(* Logix 5000 project; controller TFF vendor 1 type 14 code 107 rev 34.11; software revision 34.03; part 23 of 36 *)
(* tags used below, declared in another part *)
   Address : DINT;   // Temp Address
   Address2 : DINT;   // Temp Address
   FeedPump_PID_Settings : INT;   // Index
   Index : DINT;   // Index
   ONS_PID02 : BOOL;
   SCL : SCALE;   // Scale Instruction
   AnalogOutput : AnalogOutput[25];   // Analog Output Array
   AnalogPoint : AnalogInput[50];   // Analog Input Array
   ControlLoop : ControlLoop[20];   // Control Loop Array
   ControlLoop_FeedPump : ALIAS FOR ControlLoop[1];   // Feed Pump Control Loop
   ControlLoop_PCV001 : ALIAS FOR ControlLoop[3];   // PCV001 Control Loop
   ControlLoop_PCV001_5ms : ALIAS FOR ControlLoop[4];   // PCV001 Control Loop
   ControlLoop_PCV001_RAMP_OUT : REAL;   // Ramp Output
   ControlLoop_PCV101 : ALIAS FOR ControlLoop[5];   // PCV101 Control Loop
   Mixer : Mixer;   // Mixer config. structure
   PCV001 : ALIAS FOR AnalogPoint[3];   // Retentate Pressure Control Valve Position
   PCV001_Control : PCV_Control;   // PCV001 Control UDT
   PumpRunStatus : DINT;   // Pumps Run Status (1 = At least one pump running , 0 = no pump running)
   SIC003 : ALIAS FOR Drive[3];   // Mixer
   SIC003_AO : ALIAS FOR AnalogOutput[4];   // Mixer Speed Setpoint
   SysControl : SysControl;   // General system status and command
   WI001 : ALIAS FOR AnalogPoint[15];   // Feed Bag Weight
(* Process, continued *)

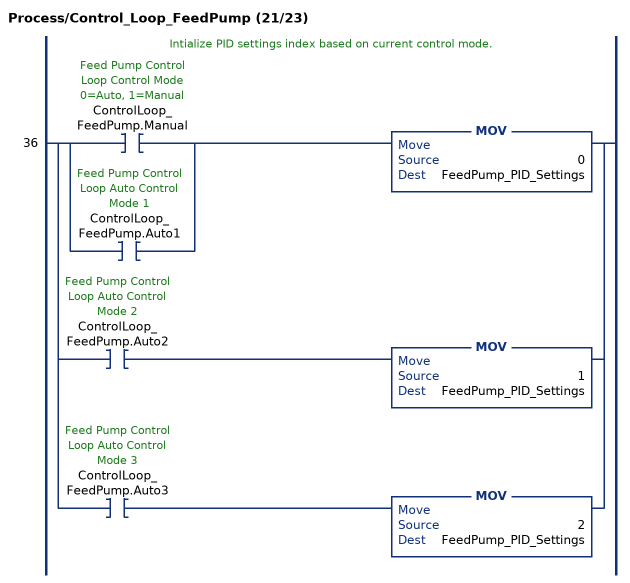
   [picture p189: Process/Control_Loop_FeedPump rungs 36-36]
   // Intialize PID settings index based on current control mode.
   36: [[XIC(ControlLoop_FeedPump.Manual) ,XIC(ControlLoop_FeedPump.Auto1) ] MOV(0,FeedPump_PID_Settings) ,XIC(ControlLoop_FeedPump.Auto2) MOV(1,FeedPump_PID_Settings) ,XIC(ControlLoop_FeedPump.Auto3) MOV(2,FeedPump_PID_Settings) ];
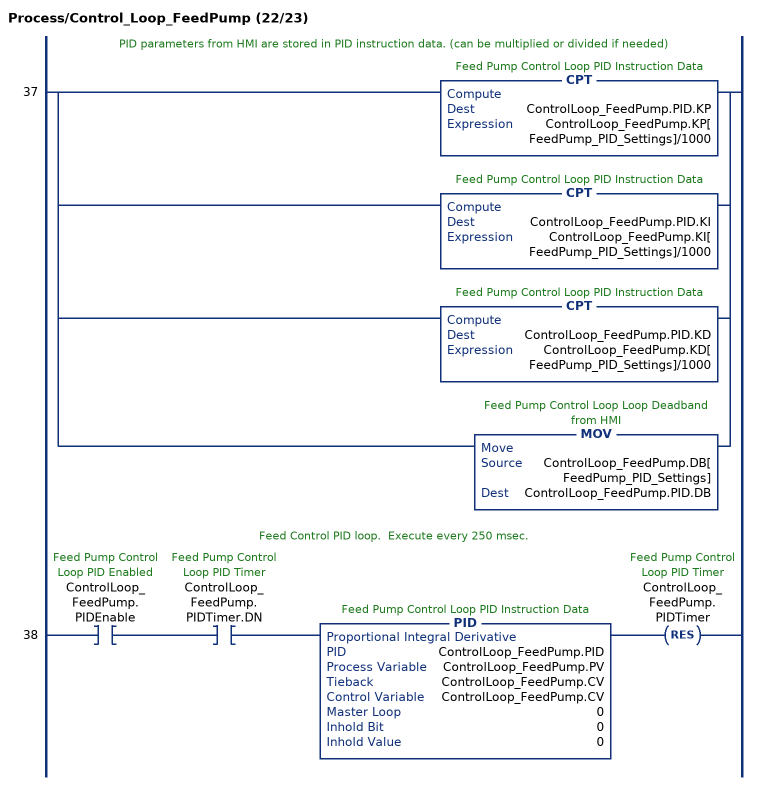
   // PID parameters from HMI are stored in PID instruction data. (can be multiplied or divided if needed)
   37: [CPT(ControlLoop_FeedPump.PID.KP,ControlLoop_FeedPump.KP[FeedPump_PID_Settings]/1000) ,CPT(ControlLoop_FeedPump.PID.KI,ControlLoop_FeedPump.KI[FeedPump_PID_Settings]/1000) ,CPT(ControlLoop_FeedPump.PID.KD,ControlLoop_FeedPump.KD[FeedPump_PID_Settings]/1000) ,MOV(ControlLoop_FeedPump.DB[FeedPump_PID_Settings],ControlLoop_FeedPump.PID.DB) ];
   // Feed Control PID loop.  Execute every 250 msec.
   38: XIC(ControlLoop_FeedPump.PIDEnable)XIC(ControlLoop_FeedPump.PIDTimer.DN)PID(ControlLoop_FeedPump.PID,ControlLoop_FeedPump.PV,ControlLoop_FeedPump.CV,ControlLoop_FeedPump.CV,0,0,0)RES(ControlLoop_FeedPump.PIDTimer);
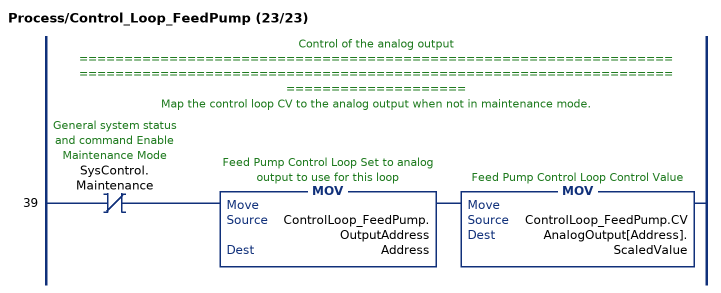
   // Control of the analog output
   // ========================================================================================================================================================
   // Map the control loop CV to the analog output when not in maintenance mode.
   39: XIO(SysControl.Maintenance)MOV(ControlLoop_FeedPump.OutputAddress,Address)MOV(ControlLoop_FeedPump.CV,AnalogOutput[Address].ScaledValue);
END_ROUTINE

ROUTINE Control_Loop_Mixer   (* ladder *)
// Agitator Control Routine
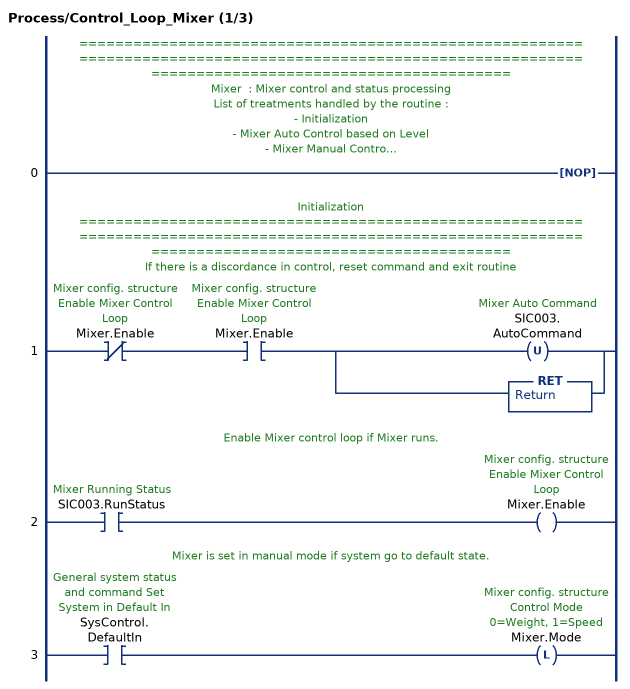
   // ========================================================================================================================================================
   //                                                                                                    Mixer  : Mixer control and status processing
   //                                                     List of treatments handled by the routine :
   //                                                          - Initialization
   //                                                          - Mixer Auto Control based on Level
   //                                                          - Mixer Manual Control
   //                                                     -----------------------------------------------------------------------------------------------------------------------------------------------------
   //                                                     History
   //                                                          2019-AUG-13 - Actemium - B. Roch - Initial version for Candidate Release 3.00.00.00.a
   // ========================================================================================================================================================
   0: NOP();
   // Initialization
   // ========================================================================================================================================================
   // If there is a discordance in control, reset command and exit routine
   1: XIO(Mixer.Enable)XIC(Mixer.Enable)[OTU(SIC003.AutoCommand) ,RET() ];
   // Enable Mixer control loop if Mixer runs.
   2: XIC(SIC003.RunStatus)OTE(Mixer.Enable);
   // Mixer is set in manual mode if system go to default state.
   3: XIC(SysControl.DefaultIn)OTL(Mixer.Mode);
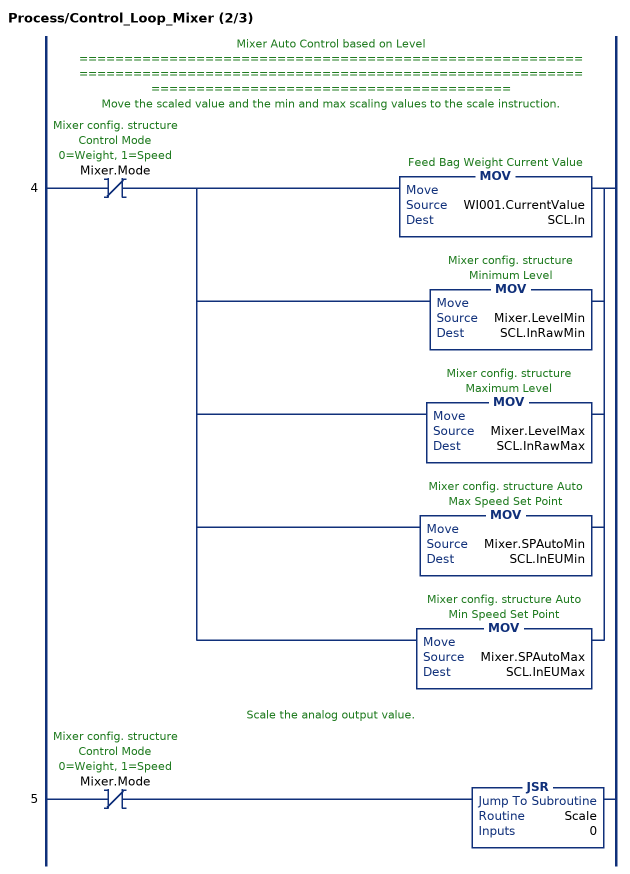
   // Mixer Auto Control based on Level
   // ========================================================================================================================================================
   // Move the scaled value and the min and max scaling values to the scale instruction.
   4: XIO(Mixer.Mode)[MOV(WI001.CurrentValue,SCL.In) ,MOV(Mixer.LevelMin,SCL.InRawMin) ,MOV(Mixer.LevelMax,SCL.InRawMax) ,MOV(Mixer.SPAutoMin,SCL.InEUMin) ,MOV(Mixer.SPAutoMax,SCL.InEUMax) ];
   // Scale the analog output value.
   5: XIO(Mixer.Mode)JSR(Scale,0);
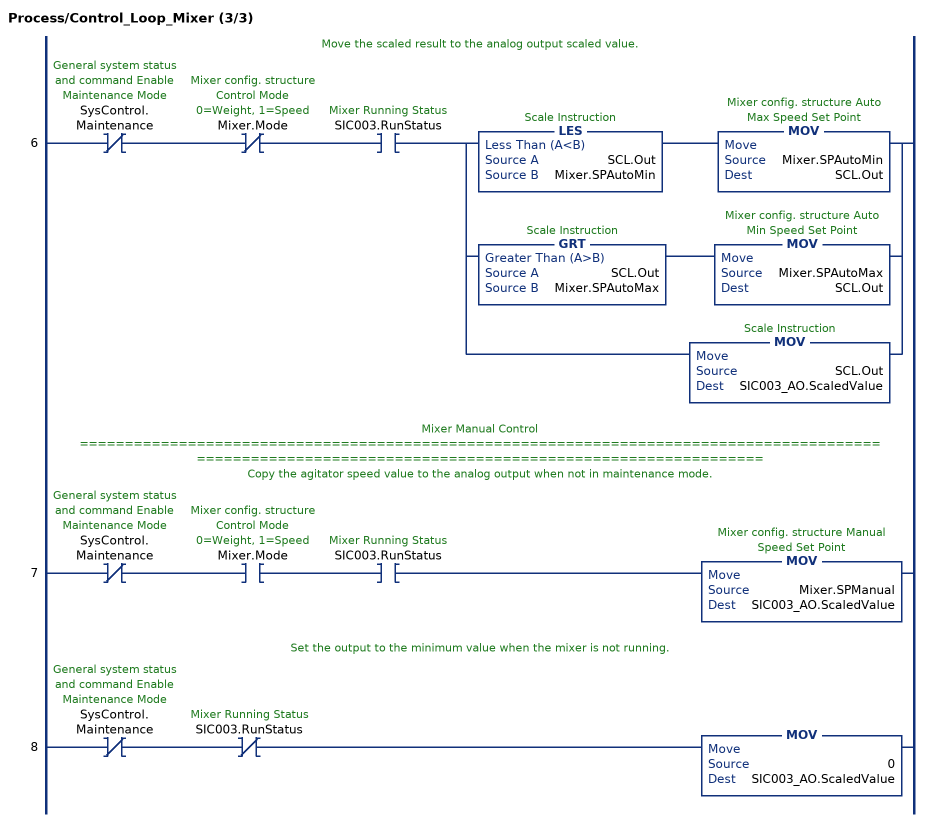
   // Move the scaled result to the analog output scaled value.
   6: XIO(SysControl.Maintenance)XIO(Mixer.Mode)XIC(SIC003.RunStatus)[LES(SCL.Out,Mixer.SPAutoMin) MOV(Mixer.SPAutoMin,SCL.Out) ,GRT(SCL.Out,Mixer.SPAutoMax) MOV(Mixer.SPAutoMax,SCL.Out) ,MOV(SCL.Out,SIC003_AO.ScaledValue) ];
   // Mixer Manual Control
   // ========================================================================================================================================================
   // Copy the agitator speed value to the analog output when not in maintenance mode.
   7: XIO(SysControl.Maintenance)XIC(Mixer.Mode)XIC(SIC003.RunStatus)MOV(Mixer.SPManual,SIC003_AO.ScaledValue);
   // Set the output to the minimum value when the mixer is not running.
   8: XIO(SysControl.Maintenance)XIO(SIC003.RunStatus)MOV(0,SIC003_AO.ScaledValue);
END_ROUTINE

ROUTINE Control_Loop_PCV001   (* ladder *)
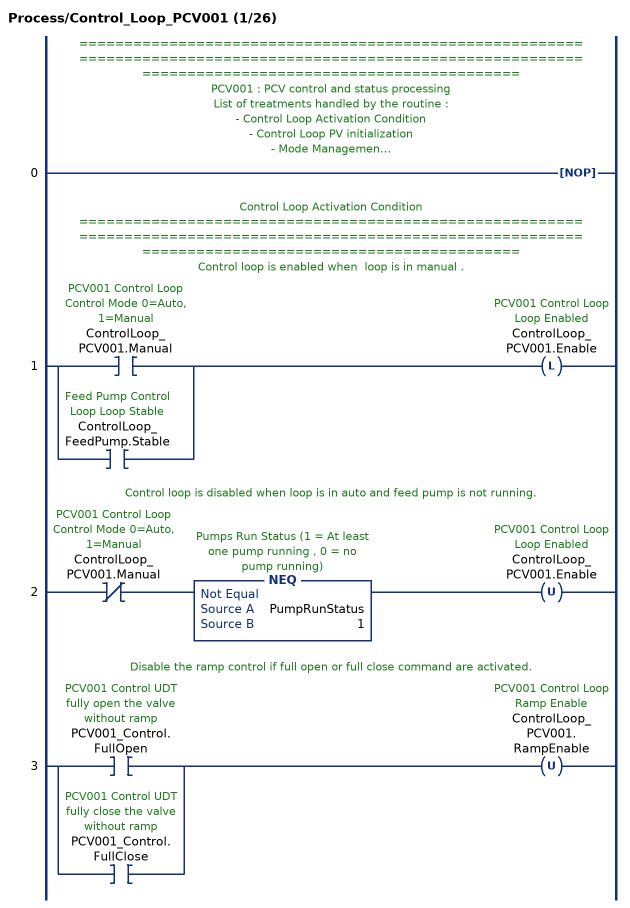
   // ==========================================================================================================================================================
   //                                                  PCV001 : PCV control and status processing
   //                                                     List of treatments handled by the routine :
   //                                                          - Control Loop Activation Condition
   //                                                  - Control Loop PV initialization
   //                                                - Mode Management
   //                                                        - Control Loop Setpoint management
   //                                                        - Control Loop deadband calculation
   //                                                          - Management of ramping control
   //                                                          - Control Loop Stability control
   //                                                          - Full Open - Full Close processing
   //                                                          - Management of PID instruction
   //                                                          - Control of the analog output
   //                                                     -----------------------------------------------------------------------------------------------------------------------------------------------------
   //                                                     History
   //                                2019-SEP-26 - Actemium - B. Roch - Initial version for Candidate Release 3.00.00.00.c                               2020-SEP-14 - Merck - Q. Spindler - Modifications for Candidate Release 3.00.00.01.a
   //                                                        - on rung 17, disable DBOK if control loop is not enabled or in manual
   // 	2021-APR-19 - DAVIDSON- Ch. ARBOGAST - Modifications for Candidate Release 3.01.00.00.a
   // 	- on rung 4, line 1, replace "ControlLoop[3].Manual OR ControlLoop[3].Auto1" by
   // 			 "NOT ControlLoop[3].Auto2 AND NOT ControlLoop[3].Auto3"
   // ==========================================================================================================================================================
   0: NOP();
   // Control Loop Activation Condition
   // ==========================================================================================================================================================
   // Control loop is enabled when  loop is in manual .
   1: [XIC(ControlLoop_PCV001.Manual) ,XIC(ControlLoop_FeedPump.Stable) ]OTL(ControlLoop_PCV001.Enable);
   // Control loop is disabled when loop is in auto and feed pump is not running.
   2: XIO(ControlLoop_PCV001.Manual)NEQ(PumpRunStatus,1)OTU(ControlLoop_PCV001.Enable);
   // Disable the ramp control if full open or full close command are activated.
   3: [XIC(PCV001_Control.FullOpen) ,XIC(PCV001_Control.FullClose) ]OTU(ControlLoop_PCV001.RampEnable);
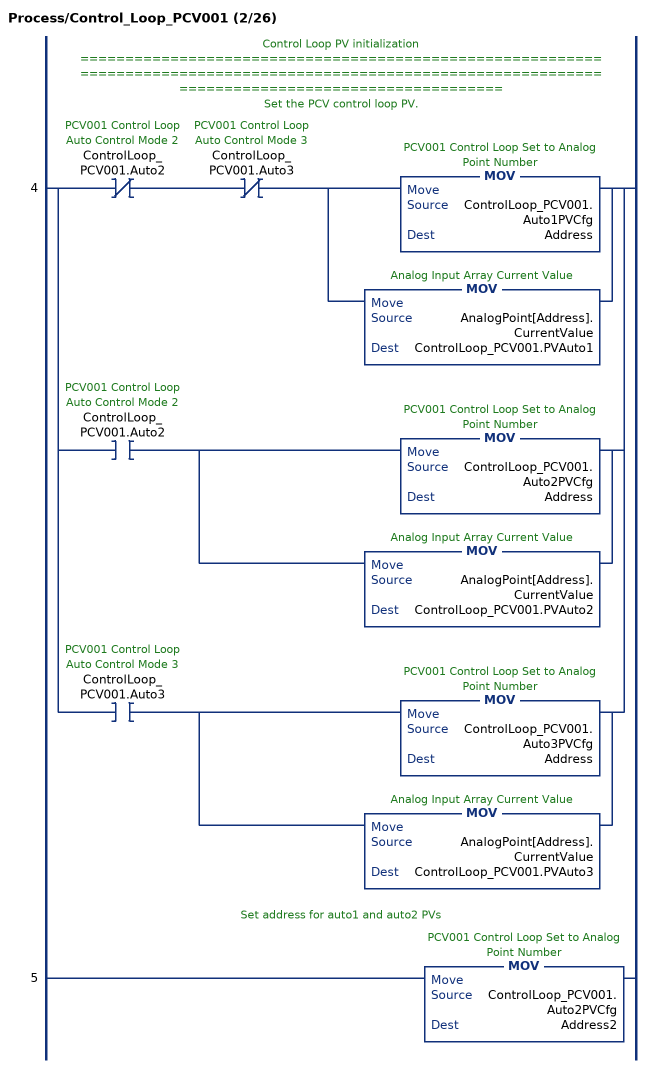
   // Control Loop PV initialization
   // ========================================================================================================================================================
   // Set the PCV control loop PV.
   4: [[XIO(ControlLoop_PCV001.Auto2) XIO(ControlLoop_PCV001.Auto3) [MOV(ControlLoop_PCV001.Auto1PVCfg,Address) ,MOV(AnalogPoint[Address].CurrentValue,ControlLoop_PCV001.PVAuto1) ] ,XIC(ControlLoop_PCV001.Auto2) [MOV(ControlLoop_PCV001.Auto2PVCfg,Address) ,MOV(AnalogPoint[Address].CurrentValue,ControlLoop_PCV001.PVAuto2) ] ] ,XIC(ControlLoop_PCV001.Auto3) [MOV(ControlLoop_PCV001.Auto3PVCfg,Address) ,MOV(AnalogPoint[Address].CurrentValue,ControlLoop_PCV001.PVAuto3) ] ];
   // Set address for auto1 and auto2 PVs
   5: MOV(ControlLoop_PCV001.Auto2PVCfg,Address2);
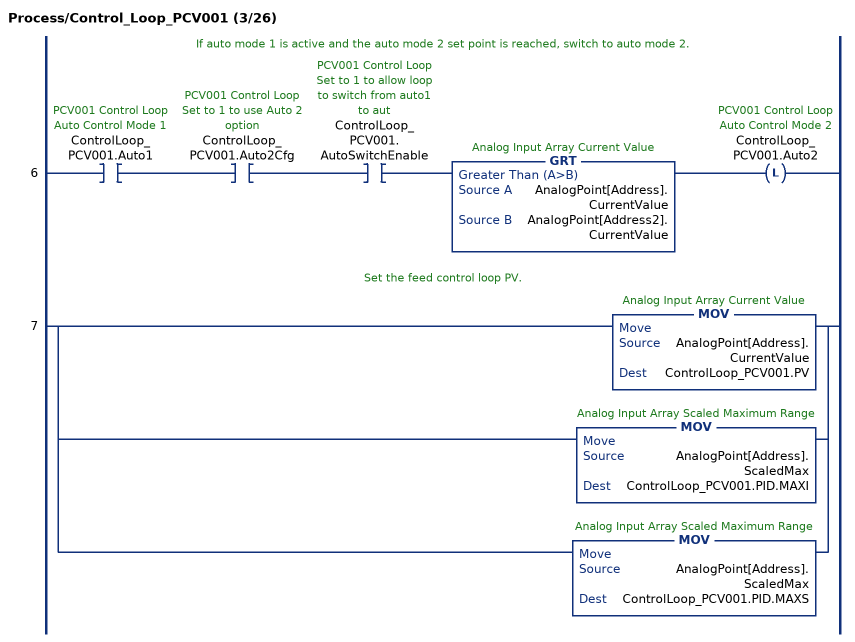
   // If auto mode 1 is active and the auto mode 2 set point is reached, switch to auto mode 2.
   6: XIC(ControlLoop_PCV001.Auto1)XIC(ControlLoop_PCV001.Auto2Cfg)XIC(ControlLoop_PCV001.AutoSwitchEnable)GRT(AnalogPoint[Address].CurrentValue,AnalogPoint[Address2].CurrentValue)OTL(ControlLoop_PCV001.Auto2);
   // Set the feed control loop PV.
   7: [MOV(AnalogPoint[Address].CurrentValue,ControlLoop_PCV001.PV) ,MOV(AnalogPoint[Address].ScaledMax,ControlLoop_PCV001.PID.MAXI) ,MOV(AnalogPoint[Address].ScaledMax,ControlLoop_PCV001.PID.MAXS) ];
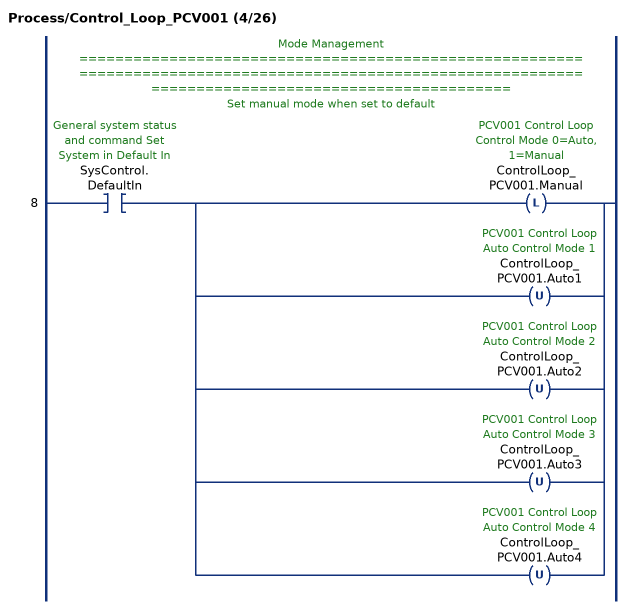
   // Mode Management
   // ========================================================================================================================================================
   // Set manual mode when set to default
   8: XIC(SysControl.DefaultIn)[OTL(ControlLoop_PCV001.Manual) ,OTU(ControlLoop_PCV001.Auto1) ,OTU(ControlLoop_PCV001.Auto2) ,OTU(ControlLoop_PCV001.Auto3) ,OTU(ControlLoop_PCV001.Auto4) ];
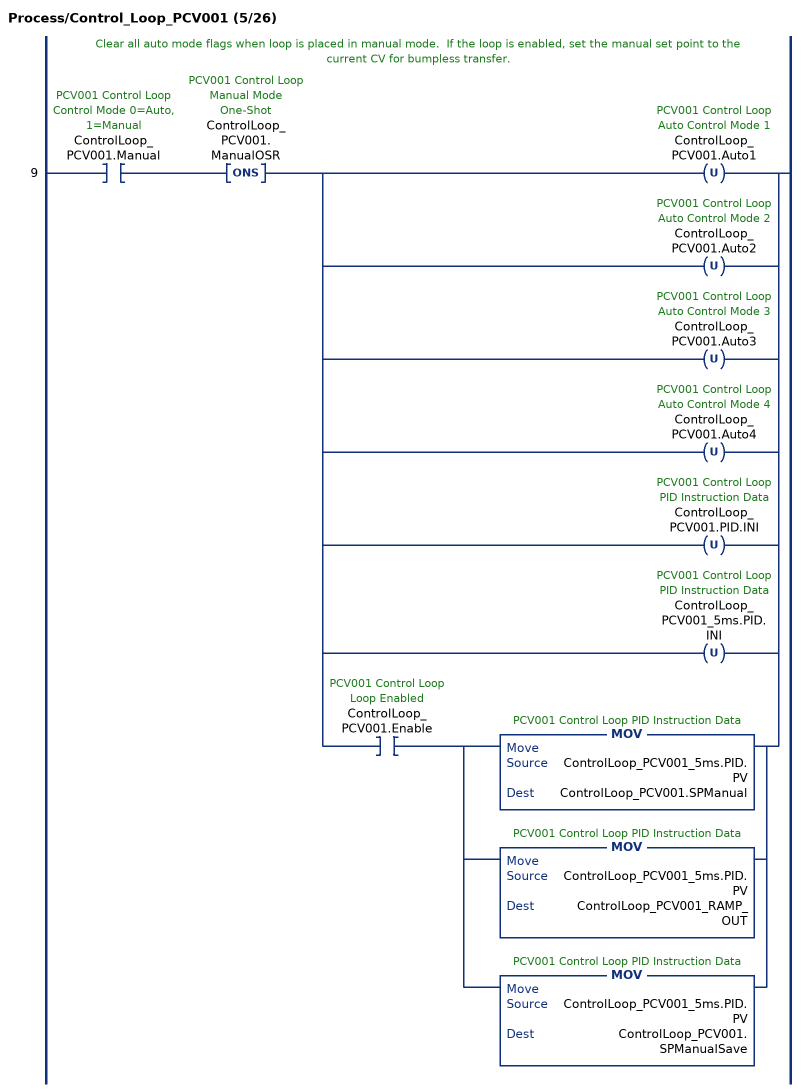
   // Clear all auto mode flags when loop is placed in manual mode.  If the loop is enabled, set the manual set point to the current CV for bumpless transfer.
   9: XIC(ControlLoop_PCV001.Manual)ONS(ControlLoop_PCV001.ManualOSR)[OTU(ControlLoop_PCV001.Auto1) ,OTU(ControlLoop_PCV001.Auto2) ,OTU(ControlLoop_PCV001.Auto3) ,OTU(ControlLoop_PCV001.Auto4) ,OTU(ControlLoop_PCV001.PID.INI) ,OTU(ControlLoop_PCV001_5ms.PID.INI) ,XIC(ControlLoop_PCV001.Enable) [MOV(ControlLoop_PCV001_5ms.PID.PV,ControlLoop_PCV001.SPManual) ,MOV(ControlLoop_PCV001_5ms.PID.PV,ControlLoop_PCV001_RAMP_OUT) ,MOV(ControlLoop_PCV001_5ms.PID.PV,ControlLoop_PCV001.SPManualSave) ] ];
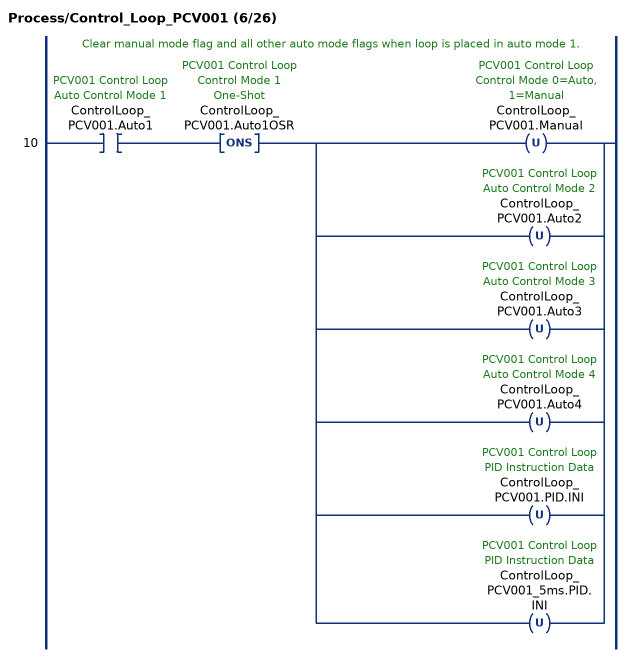
   // Clear manual mode flag and all other auto mode flags when loop is placed in auto mode 1.
   10: XIC(ControlLoop_PCV001.Auto1)ONS(ControlLoop_PCV001.Auto1OSR)[OTU(ControlLoop_PCV001.Manual) ,OTU(ControlLoop_PCV001.Auto2) ,OTU(ControlLoop_PCV001.Auto3) ,OTU(ControlLoop_PCV001.Auto4) ,OTU(ControlLoop_PCV001.PID.INI) ,OTU(ControlLoop_PCV001_5ms.PID.INI) ];
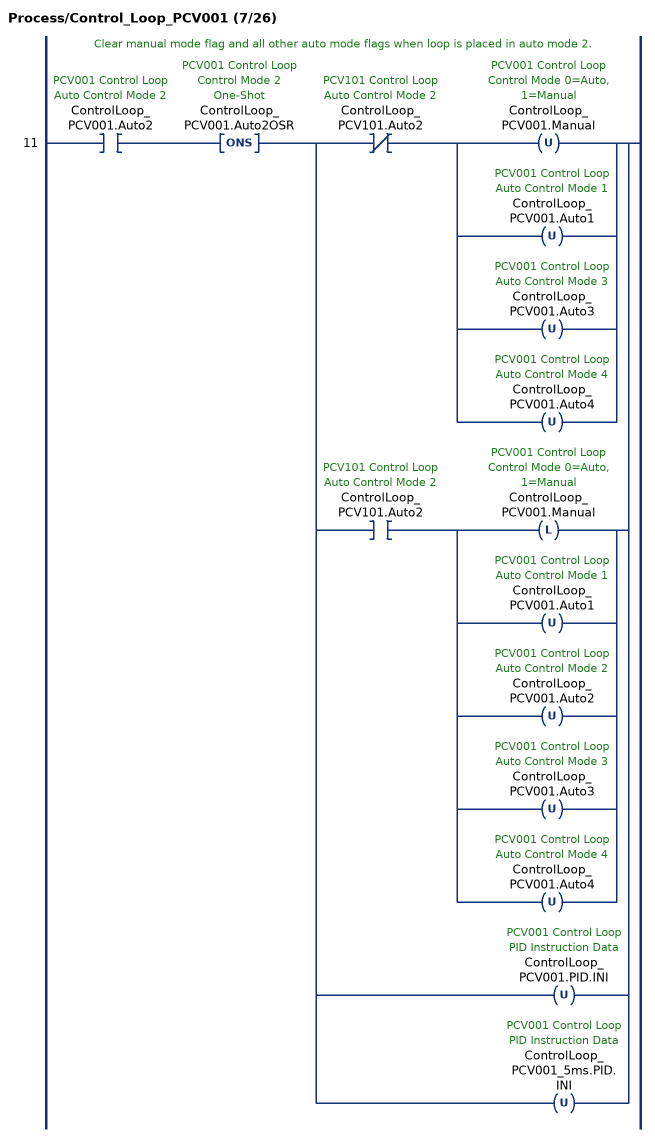
   // Clear manual mode flag and all other auto mode flags when loop is placed in auto mode 2.
   11: XIC(ControlLoop_PCV001.Auto2)ONS(ControlLoop_PCV001.Auto2OSR)[XIO(ControlLoop_PCV101.Auto2) [OTU(ControlLoop_PCV001.Manual) ,OTU(ControlLoop_PCV001.Auto1) ,OTU(ControlLoop_PCV001.Auto3) ,OTU(ControlLoop_PCV001.Auto4) ] ,XIC(ControlLoop_PCV101.Auto2) [OTL(ControlLoop_PCV001.Manual) ,OTU(ControlLoop_PCV001.Auto1) ,OTU(ControlLoop_PCV001.Auto2) ,OTU(ControlLoop_PCV001.Auto3) ,OTU(ControlLoop_PCV001.Auto4) ] ,OTU(ControlLoop_PCV001.PID.INI) ,OTU(ControlLoop_PCV001_5ms.PID.INI) ];
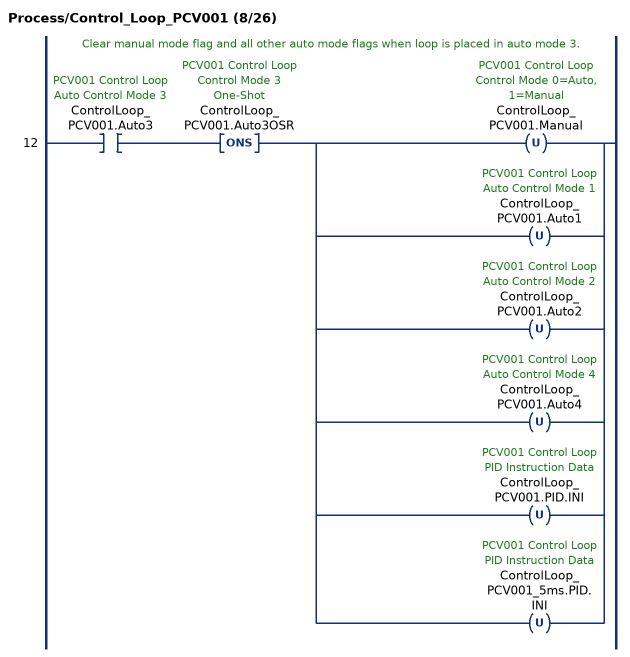
   // Clear manual mode flag and all other auto mode flags when loop is placed in auto mode 3.
   12: XIC(ControlLoop_PCV001.Auto3)ONS(ControlLoop_PCV001.Auto3OSR)[OTU(ControlLoop_PCV001.Manual) ,OTU(ControlLoop_PCV001.Auto1) ,OTU(ControlLoop_PCV001.Auto2) ,OTU(ControlLoop_PCV001.Auto4) ,OTU(ControlLoop_PCV001.PID.INI) ,OTU(ControlLoop_PCV001_5ms.PID.INI) ];
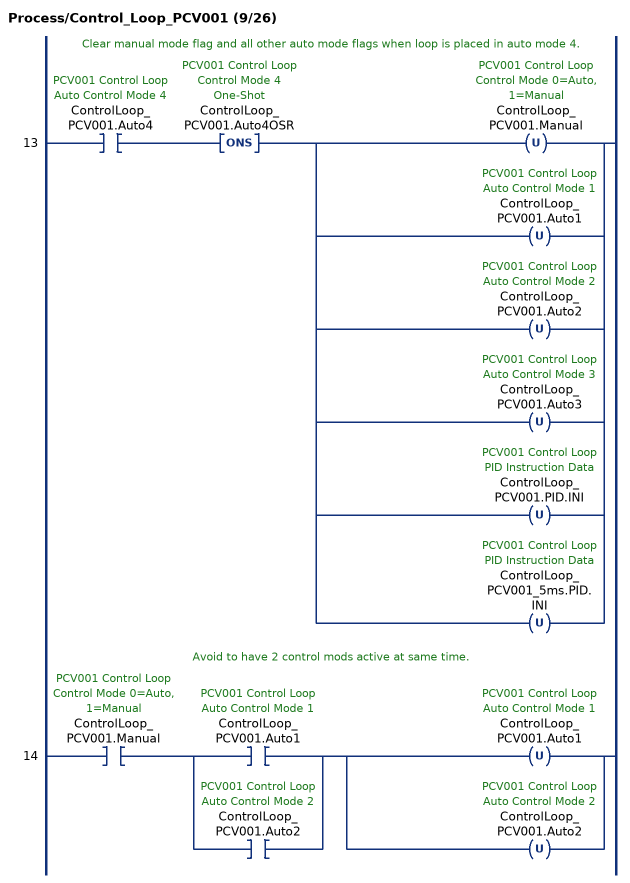
   // Clear manual mode flag and all other auto mode flags when loop is placed in auto mode 4.
   13: XIC(ControlLoop_PCV001.Auto4)ONS(ControlLoop_PCV001.Auto4OSR)[OTU(ControlLoop_PCV001.Manual) ,OTU(ControlLoop_PCV001.Auto1) ,OTU(ControlLoop_PCV001.Auto2) ,OTU(ControlLoop_PCV001.Auto3) ,OTU(ControlLoop_PCV001.PID.INI) ,OTU(ControlLoop_PCV001_5ms.PID.INI) ];
   // Avoid to have 2 control mods active at same time.
   14: XIC(ControlLoop_PCV001.Manual)[XIC(ControlLoop_PCV001.Auto1) ,XIC(ControlLoop_PCV001.Auto2) ][OTU(ControlLoop_PCV001.Auto1) ,OTU(ControlLoop_PCV001.Auto2) ];
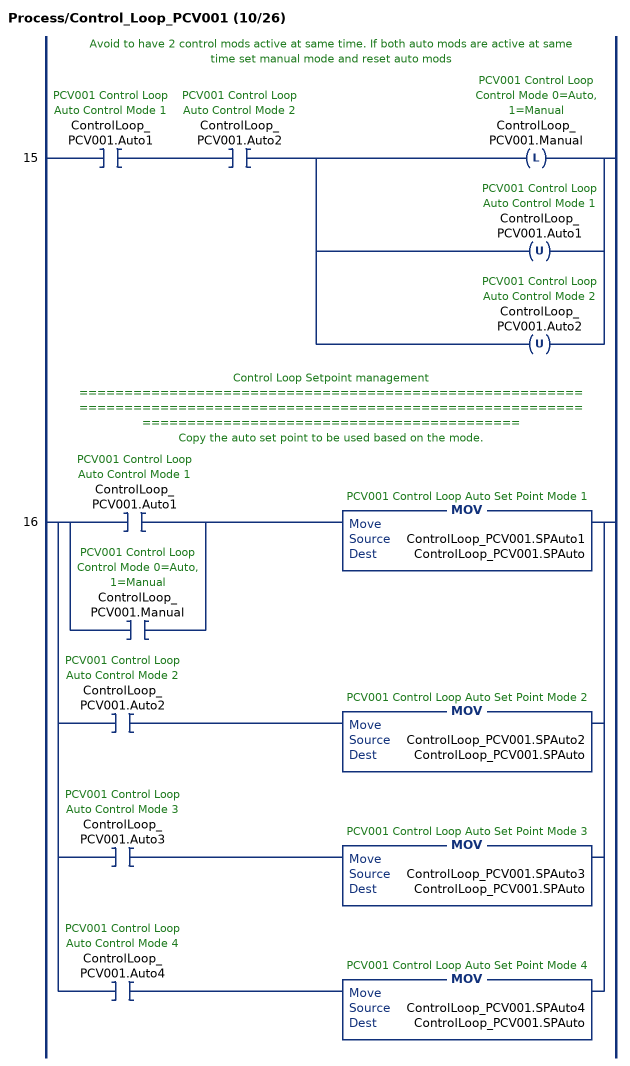
   // Avoid to have 2 control mods active at same time. If both auto mods are active at same time set manual mode and reset auto mods
   15: XIC(ControlLoop_PCV001.Auto1)XIC(ControlLoop_PCV001.Auto2)[OTL(ControlLoop_PCV001.Manual) ,OTU(ControlLoop_PCV001.Auto1) ,OTU(ControlLoop_PCV001.Auto2) ];
   // Control Loop Setpoint management
   // ==========================================================================================================================================================
   // Copy the auto set point to be used based on the mode.
   16: [[XIC(ControlLoop_PCV001.Auto1) ,XIC(ControlLoop_PCV001.Manual) ] MOV(ControlLoop_PCV001.SPAuto1,ControlLoop_PCV001.SPAuto) ,XIC(ControlLoop_PCV001.Auto2) MOV(ControlLoop_PCV001.SPAuto2,ControlLoop_PCV001.SPAuto) ,XIC(ControlLoop_PCV001.Auto3) MOV(ControlLoop_PCV001.SPAuto3,ControlLoop_PCV001.SPAuto) ,XIC(ControlLoop_PCV001.Auto4) MOV(ControlLoop_PCV001.SPAuto4,ControlLoop_PCV001.SPAuto) ];
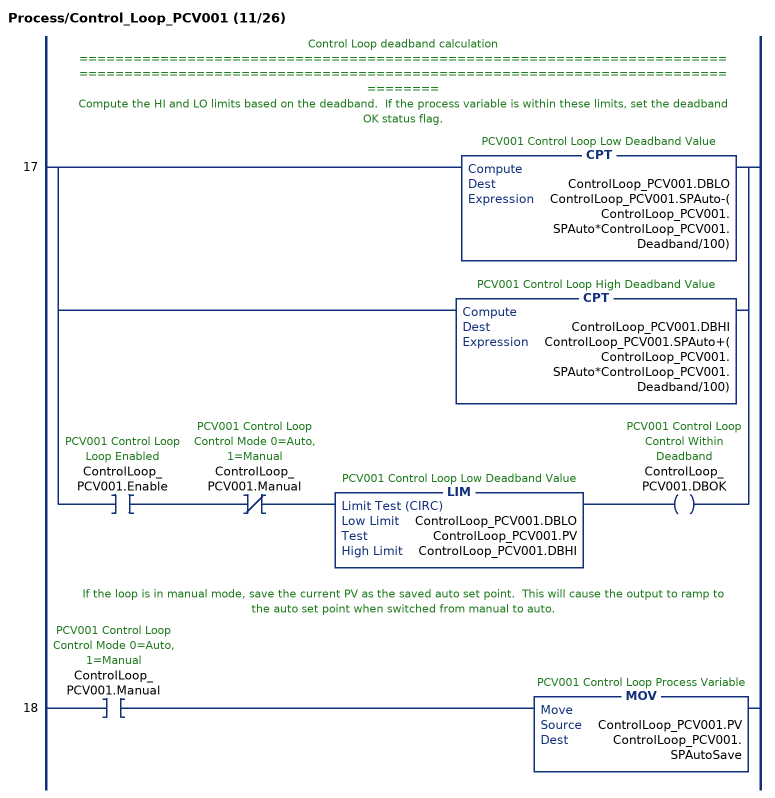
   // Control Loop deadband calculation
   // ========================================================================================================================================================
   // Compute the HI and LO limits based on the deadband.  If the process variable is within these limits, set the deadband OK status flag.
   17: [CPT(ControlLoop_PCV001.DBLO,ControlLoop_PCV001.SPAuto-(ControlLoop_PCV001.SPAuto*ControlLoop_PCV001.Deadband/100)) ,CPT(ControlLoop_PCV001.DBHI,ControlLoop_PCV001.SPAuto+(ControlLoop_PCV001.SPAuto*ControlLoop_PCV001.Deadband/100)) ,XIC(ControlLoop_PCV001.Enable) XIO(ControlLoop_PCV001.Manual) LIM(ControlLoop_PCV001.DBLO,ControlLoop_PCV001.PV,ControlLoop_PCV001.DBHI) OTE(ControlLoop_PCV001.DBOK) ];
   // If the loop is in manual mode, save the current PV as the saved auto set point.  This will cause the output to ramp to the auto set point when switched from manual to auto.
   18: XIC(ControlLoop_PCV001.Manual)MOV(ControlLoop_PCV001.PV,ControlLoop_PCV001.SPAutoSave);
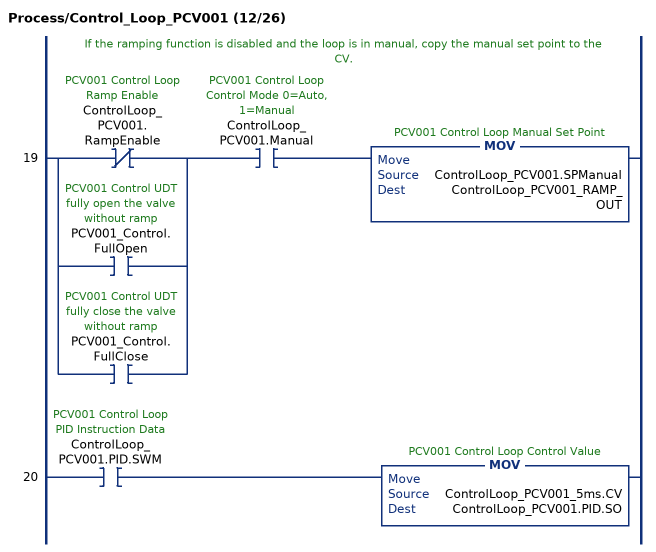
   // If the ramping function is disabled and the loop is in manual, copy the manual set point to the CV.
   19: [XIO(ControlLoop_PCV001.RampEnable) ,XIC(PCV001_Control.FullOpen) ,XIC(PCV001_Control.FullClose) ]XIC(ControlLoop_PCV001.Manual)MOV(ControlLoop_PCV001.SPManual,ControlLoop_PCV001_RAMP_OUT);
   20: XIC(ControlLoop_PCV001.PID.SWM)MOV(ControlLoop_PCV001_5ms.CV,ControlLoop_PCV001.PID.SO);
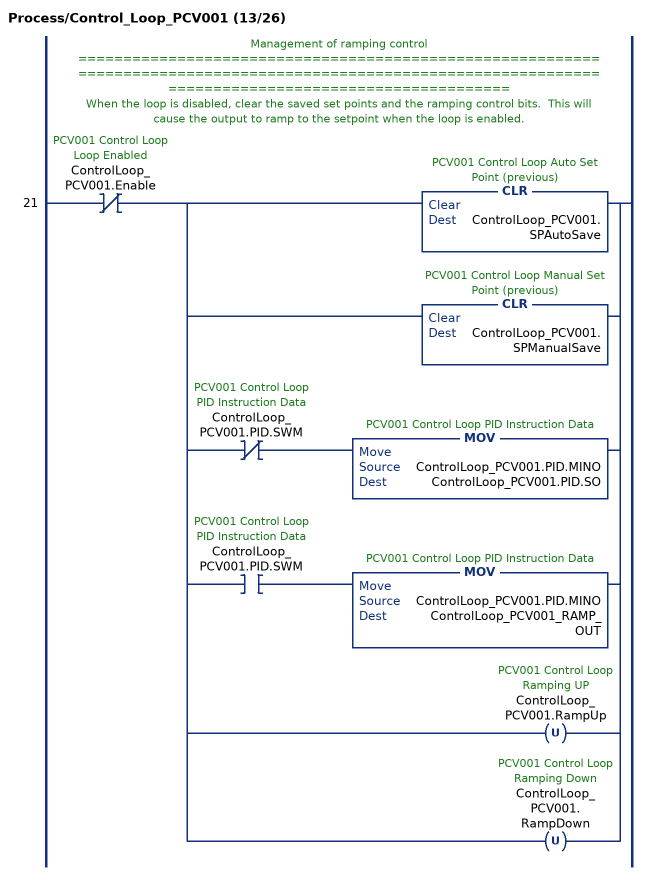
   // Management of ramping control
   // ==========================================================================================================================================================
   // When the loop is disabled, clear the saved set points and the ramping control bits.  This will cause the output to ramp to the setpoint when the loop is enabled.
   21: XIO(ControlLoop_PCV001.Enable)[CLR(ControlLoop_PCV001.SPAutoSave) ,CLR(ControlLoop_PCV001.SPManualSave) ,XIO(ControlLoop_PCV001.PID.SWM) MOV(ControlLoop_PCV001.PID.MINO,ControlLoop_PCV001.PID.SO) ,XIC(ControlLoop_PCV001.PID.SWM) MOV(ControlLoop_PCV001.PID.MINO,ControlLoop_PCV001_RAMP_OUT) ,OTU(ControlLoop_PCV001.RampUp) ,OTU(ControlLoop_PCV001.RampDown) ];
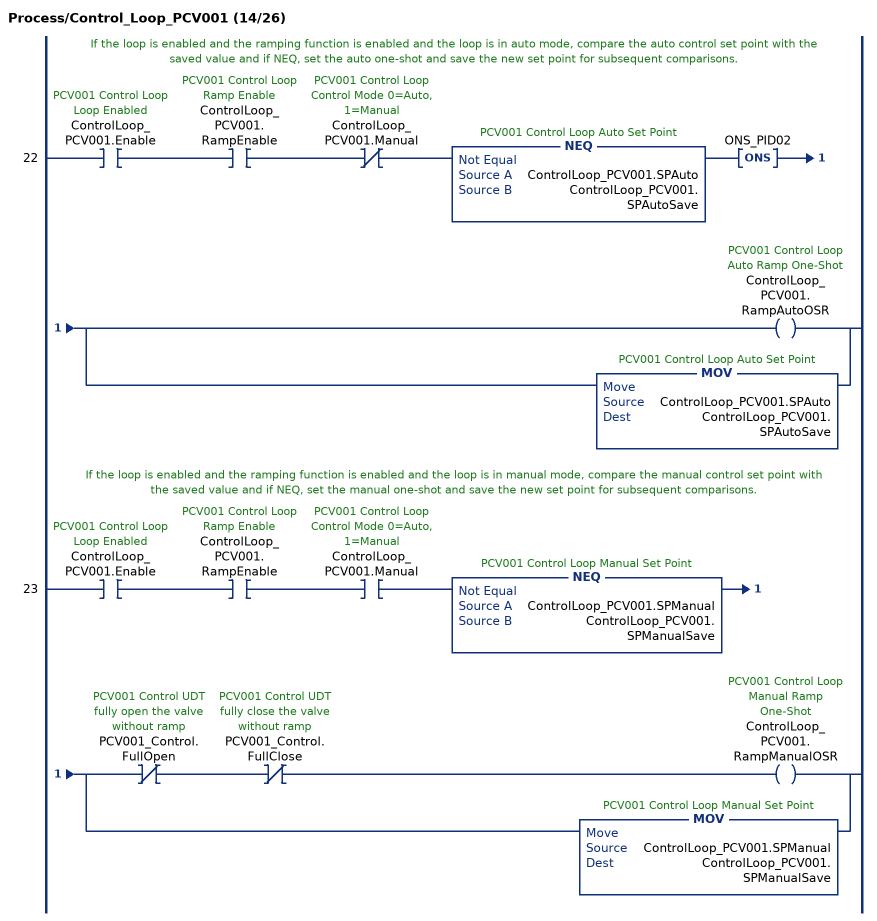
   // If the loop is enabled and the ramping function is enabled and the loop is in auto mode, compare the auto control set point with the saved value and if NEQ, set the auto one-shot and save the new set point for subsequent comparisons.
   22: XIC(ControlLoop_PCV001.Enable)XIC(ControlLoop_PCV001.RampEnable)XIO(ControlLoop_PCV001.Manual)NEQ(ControlLoop_PCV001.SPAuto,ControlLoop_PCV001.SPAutoSave)ONS(ONS_PID02)[OTE(ControlLoop_PCV001.RampAutoOSR) ,MOV(ControlLoop_PCV001.SPAuto,ControlLoop_PCV001.SPAutoSave) ];
   // If the loop is enabled and the ramping function is enabled and the loop is in manual mode, compare the manual control set point with the saved value and if NEQ, set the manual one-shot and save the new set point for subsequent comparisons.
   23: XIC(ControlLoop_PCV001.Enable)XIC(ControlLoop_PCV001.RampEnable)XIC(ControlLoop_PCV001.Manual)NEQ(ControlLoop_PCV001.SPManual,ControlLoop_PCV001.SPManualSave)[XIO(PCV001_Control.FullOpen) XIO(PCV001_Control.FullClose) OTE(ControlLoop_PCV001.RampManualOSR) ,MOV(ControlLoop_PCV001.SPManual,ControlLoop_PCV001.SPManualSave) ];
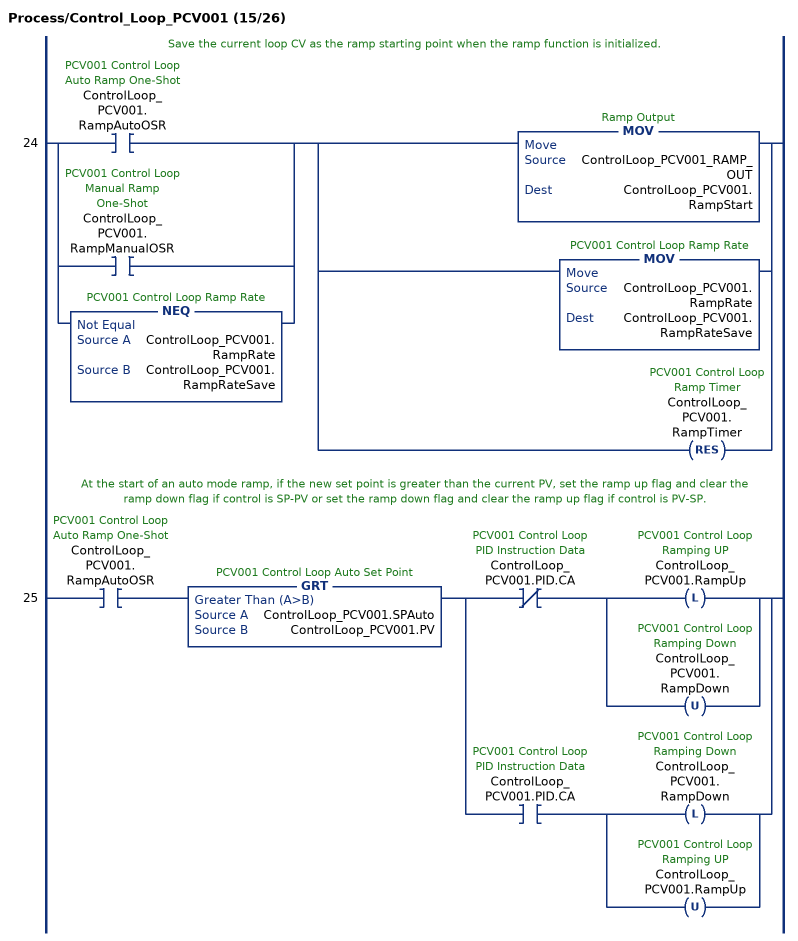
   // Save the current loop CV as the ramp starting point when the ramp function is initialized.
   24: [XIC(ControlLoop_PCV001.RampAutoOSR) ,XIC(ControlLoop_PCV001.RampManualOSR) ,NEQ(ControlLoop_PCV001.RampRate,ControlLoop_PCV001.RampRateSave) ][MOV(ControlLoop_PCV001_RAMP_OUT,ControlLoop_PCV001.RampStart) ,MOV(ControlLoop_PCV001.RampRate,ControlLoop_PCV001.RampRateSave) ,RES(ControlLoop_PCV001.RampTimer) ];
   // At the start of an auto mode ramp, if the new set point is greater than the current PV, set the ramp up flag and clear the ramp down flag if control is SP-PV or set the ramp down flag and clear the ramp up flag if control is PV-SP.
   25: XIC(ControlLoop_PCV001.RampAutoOSR)GRT(ControlLoop_PCV001.SPAuto,ControlLoop_PCV001.PV)[XIO(ControlLoop_PCV001.PID.CA) [OTL(ControlLoop_PCV001.RampUp) ,OTU(ControlLoop_PCV001.RampDown) ] ,XIC(ControlLoop_PCV001.PID.CA) [OTL(ControlLoop_PCV001.RampDown) ,OTU(ControlLoop_PCV001.RampUp) ] ];
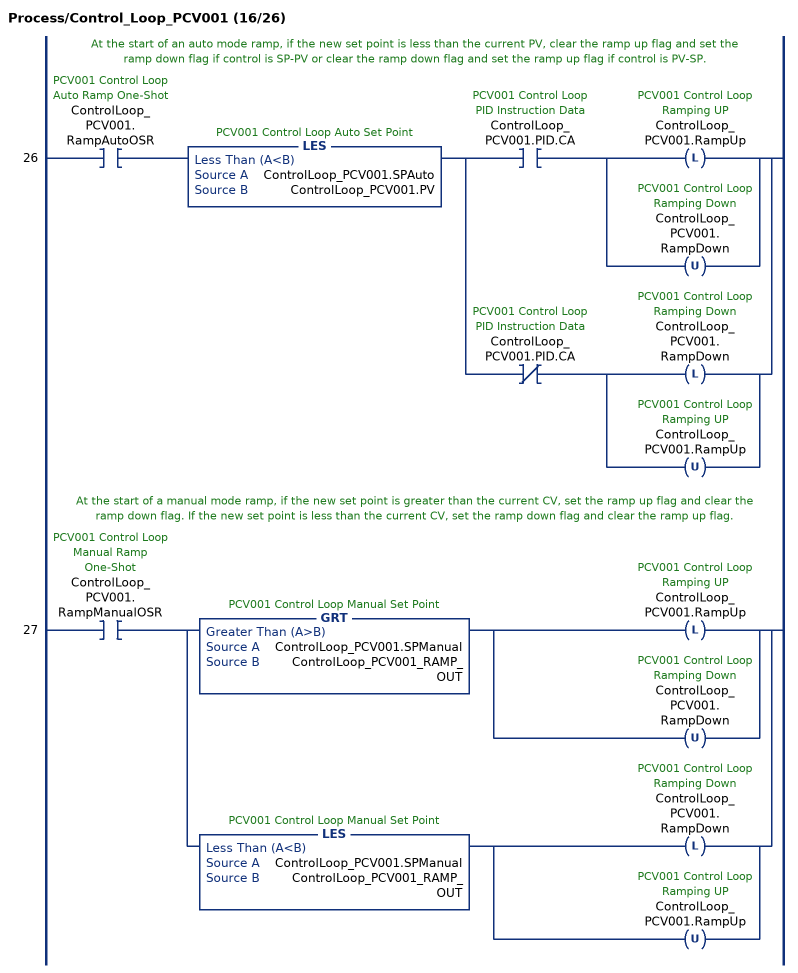
   // At the start of an auto mode ramp, if the new set point is less than the current PV, clear the ramp up flag and set the ramp down flag if control is SP-PV or clear the ramp down flag and set the ramp up flag if control is PV-SP.
   26: XIC(ControlLoop_PCV001.RampAutoOSR)LES(ControlLoop_PCV001.SPAuto,ControlLoop_PCV001.PV)[XIC(ControlLoop_PCV001.PID.CA) [OTL(ControlLoop_PCV001.RampUp) ,OTU(ControlLoop_PCV001.RampDown) ] ,XIO(ControlLoop_PCV001.PID.CA) [OTL(ControlLoop_PCV001.RampDown) ,OTU(ControlLoop_PCV001.RampUp) ] ];
   // At the start of a manual mode ramp, if the new set point is greater than the current CV, set the ramp up flag and clear the ramp down flag. If the new set point is less than the current CV, set the ramp down flag and clear the ramp up flag.
   27: XIC(ControlLoop_PCV001.RampManualOSR)[GRT(ControlLoop_PCV001.SPManual,ControlLoop_PCV001_RAMP_OUT) [OTL(ControlLoop_PCV001.RampUp) ,OTU(ControlLoop_PCV001.RampDown) ] ,LES(ControlLoop_PCV001.SPManual,ControlLoop_PCV001_RAMP_OUT) [OTL(ControlLoop_PCV001.RampDown) ,OTU(ControlLoop_PCV001.RampUp) ] ];
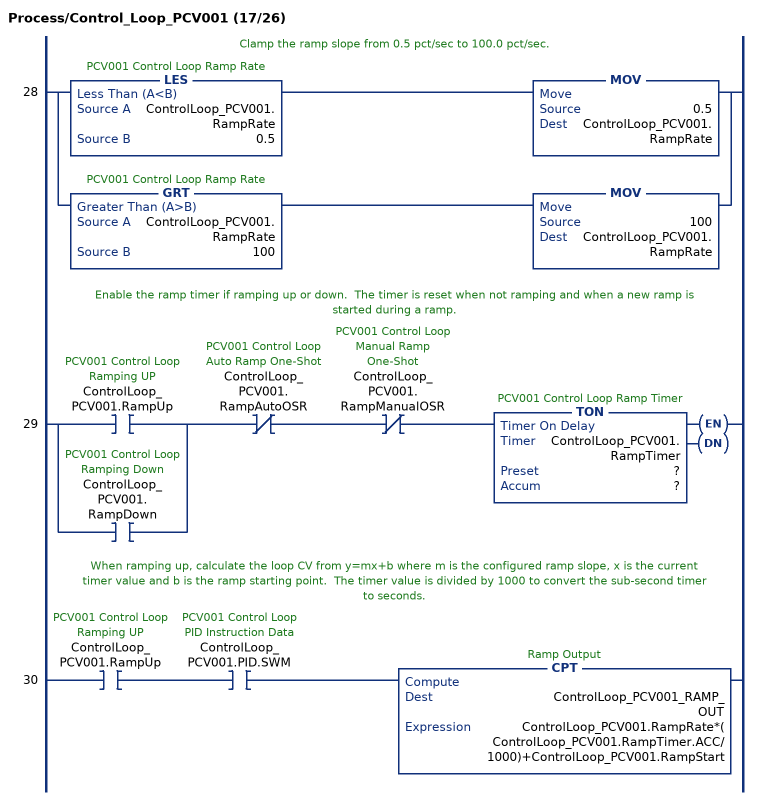
   // Clamp the ramp slope from 0.5 pct/sec to 100.0 pct/sec.
   28: [LES(ControlLoop_PCV001.RampRate,0.5) MOV(0.5,ControlLoop_PCV001.RampRate) ,GRT(ControlLoop_PCV001.RampRate,100) MOV(100,ControlLoop_PCV001.RampRate) ];
   // Enable the ramp timer if ramping up or down.  The timer is reset when not ramping and when a new ramp is started during a ramp.
   29: [XIC(ControlLoop_PCV001.RampUp) ,XIC(ControlLoop_PCV001.RampDown) ]XIO(ControlLoop_PCV001.RampAutoOSR)XIO(ControlLoop_PCV001.RampManualOSR)TON(ControlLoop_PCV001.RampTimer,?,?);
   // When ramping up, calculate the loop CV from y=mx+b where m is the configured ramp slope, x is the current timer value and b is the ramp starting point.  The timer value is divided by 1000 to convert the sub-second timer to seconds.
   30: XIC(ControlLoop_PCV001.RampUp)XIC(ControlLoop_PCV001.PID.SWM)CPT(ControlLoop_PCV001_RAMP_OUT,ControlLoop_PCV001.RampRate*(ControlLoop_PCV001.RampTimer.ACC/1000)+ControlLoop_PCV001.RampStart);
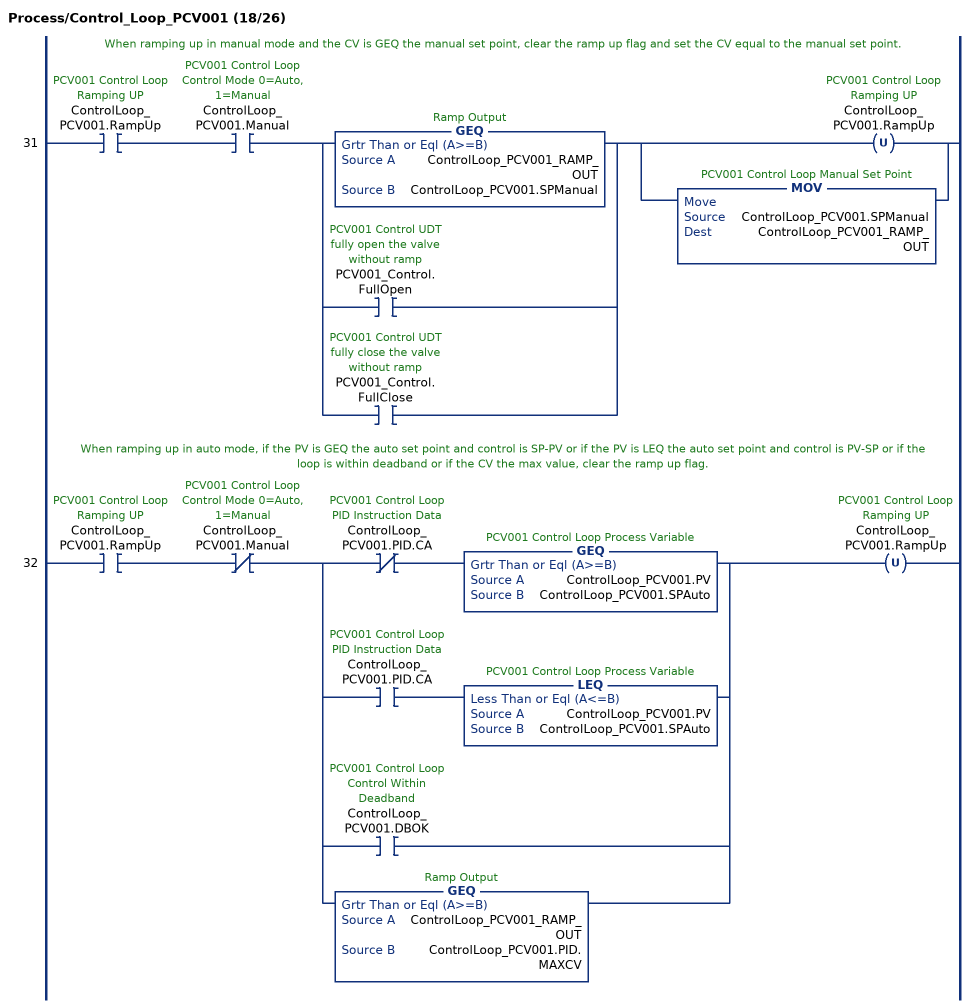
   // When ramping up in manual mode and the CV is GEQ the manual set point, clear the ramp up flag and set the CV equal to the manual set point.
   31: XIC(ControlLoop_PCV001.RampUp)XIC(ControlLoop_PCV001.Manual)[GEQ(ControlLoop_PCV001_RAMP_OUT,ControlLoop_PCV001.SPManual) ,XIC(PCV001_Control.FullOpen) ,XIC(PCV001_Control.FullClose) ][OTU(ControlLoop_PCV001.RampUp) ,MOV(ControlLoop_PCV001.SPManual,ControlLoop_PCV001_RAMP_OUT) ];
   // When ramping up in auto mode, if the PV is GEQ the auto set point and control is SP-PV or if the PV is LEQ the auto set point and control is PV-SP or if the loop is within deadband or if the CV the max value, clear the ramp up flag.
   32: XIC(ControlLoop_PCV001.RampUp)XIO(ControlLoop_PCV001.Manual)[XIO(ControlLoop_PCV001.PID.CA) GEQ(ControlLoop_PCV001.PV,ControlLoop_PCV001.SPAuto) ,XIC(ControlLoop_PCV001.PID.CA) LEQ(ControlLoop_PCV001.PV,ControlLoop_PCV001.SPAuto) ,XIC(ControlLoop_PCV001.DBOK) ,GEQ(ControlLoop_PCV001_RAMP_OUT,ControlLoop_PCV001.PID.MAXCV) ]OTU(ControlLoop_PCV001.RampUp);
